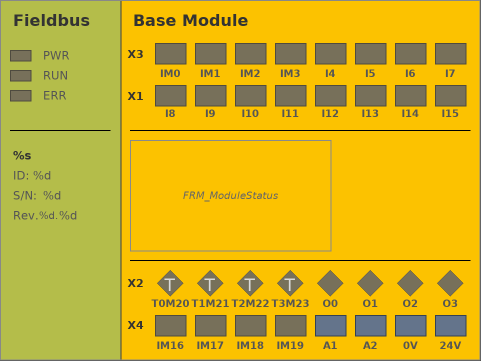
VISUALIZATION FRM_ModuleBase  // 481x361
VAR_IN_OUT
   stFieldbusData: ST_PNOZModuleData;
   stBaseModuleData: ST_PNOZModuleData;
END_VAR
    Rectangle (120,0 361x361)
    Frame (130,140 201x111)
        shows FRM_ModuleStatus(bPower := stBaseModuleData.stLEDState.bPower, bRun := stBaseModuleData.stLEDState.bRun, bDiag := stBaseModuleData.stLEDState.bDiag, bFault := stBaseModuleData.stLEDState.bFault, bInputFault := stBaseModuleData.stLEDState.bInputFault, bOutputFault := stBaseModuleData.stLEDState.bOutputFault, sName := stBaseModuleData.sName, nID := stBaseModuleData.nID, nSerialNumber := stBaseModuleData.nSerialNumber, anRevision := stBaseModuleData.anDeviceVersion)
    Line (130,130) (470,130)
    Line (130,260) (470,260)
    Label (120,44 31x21), "X3"
    Label (120,86 31x21), "X1"
    Label (120,273 31x21), "X2"
    Label (120,315 31x21), "X4"
    Label (130,0 141x41), "Base Module"
    Rectangle (0,0 121x361)
    Label (10,0 101x41), "Fieldbus"
    Rectangle (10,50 21x11), colour toggle: stFieldbusData.stLEDState.bPower
    Label (40,50 41x11), "PWR"
    Rectangle (10,70 21x11), colour toggle: stFieldbusData.stLEDState.bRun
    Label (40,70 41x11), "RUN"
    Rectangle (10,90 21x11), colour toggle: stFieldbusData.stLEDState.bFault
    Label (40,90 41x11), "ERR"
    Textfield (40,190 71x11), "%d", text variable: stFieldbusData.nSerialNumber
    Textfield (30,170 81x11), "%d", text variable: stFieldbusData.nID
    Textfield (10,150 101x11), "%s", text variable: stFieldbusData.sName
    Label (10,170 21x11), "ID:"
    Label (10,190 31x11), "S/N:"
    Line (10,130) (110,130)
    Rectangle (155,43 31x21), colour toggle: stBaseModuleData.anInput[1].b0
    Rectangle (195,43 31x21), colour toggle: stBaseModuleData.anInput[1].b1
    Rectangle (235,43 31x21), colour toggle: stBaseModuleData.anInput[1].b2
    Rectangle (275,43 31x21), colour toggle: stBaseModuleData.anInput[1].b3
    Rectangle (315,43 31x21), colour toggle: stBaseModuleData.anInput[1].b4
    Rectangle (355,43 31x21), colour toggle: stBaseModuleData.anInput[1].b5
    Rectangle (395,43 31x21), colour toggle: stBaseModuleData.anInput[1].b6
    Rectangle (435,43 31x21), colour toggle: stBaseModuleData.anInput[1].b7
    Label (150,68 41x11), "IM0"
    Label (190,68 41x11), "IM1"
    Label (230,68 41x11), "IM2"
    Label (270,68 41x11), "IM3"
    Label (310,68 41x11), "I4"
    Label (350,68 41x11), "I5"
    Label (390,68 41x11), "I6"
    Label (430,68 41x11), "I7"
    Rectangle (155,85 31x21), colour toggle: stBaseModuleData.anInput[2].b0
    Label (150,108 41x11), "I8"
    Label (190,108 41x11), "I9"
    Label (230,108 41x11), "I10"
    Label (270,108 41x11), "I11"
    Label (310,108 41x11), "I12"
    Label (350,108 41x11), "I13"
    Label (390,108 41x11), "I14"
    Label (430,108 41x11), "I15"
    Rectangle (195,85 31x21), colour toggle: stBaseModuleData.anInput[2].b1
    Rectangle (235,85 31x21), colour toggle: stBaseModuleData.anInput[2].b2
    Rectangle (275,85 31x21), colour toggle: stBaseModuleData.anInput[2].b3
    Rectangle (315,85 31x21), colour toggle: stBaseModuleData.anInput[2].b3
    Rectangle (355,85 31x21), colour toggle: stBaseModuleData.anInput[2].b5
    Rectangle (395,85 31x21), colour toggle: stBaseModuleData.anInput[2].b6
    Rectangle (435,85 31x21), colour toggle: stBaseModuleData.anInput[2].b7
    Polygon (157,283) (170,270) (183,283) (170,296) (170,296), colour toggle: stBaseModuleData.anOutput[2].b4
    Label (150,298 41x11), "T0M20"
    Label (190,298 41x11), "T1M21"
    Label (230,298 41x11), "T2M22"
    Label (270,298 41x11), "T3M23"
    Label (310,298 41x11), "O0"
    Label (350,298 41x11), "O1"
    Label (390,298 41x11), "O2"
    Label (430,298 41x11), "O3"
    Polygon (197,283) (210,270) (223,283) (210,296) (210,296), colour toggle: stBaseModuleData.anOutput[2].b5
    Polygon (237,283) (250,270) (263,283) (250,296) (250,296), colour toggle: stBaseModuleData.anOutput[2].b6
    Polygon (277,283) (290,270) (303,283) (290,296) (290,296), colour toggle: stBaseModuleData.anOutput[2].b7
    Polygon (317,283) (330,270) (343,283) (330,296) (330,296), colour toggle: stBaseModuleData.anOutput[1].b0
    Polygon (357,283) (370,270) (383,283) (370,296) (370,296), colour toggle: stBaseModuleData.anOutput[1].b1
    Polygon (397,283) (410,270) (423,283) (410,296) (410,296), colour toggle: stBaseModuleData.anOutput[1].b2
    Polygon (437,283) (450,270) (463,283) (450,296) (450,296), colour toggle: stBaseModuleData.anOutput[1].b3
    Rectangle (155,315 31x21), colour toggle: stBaseModuleData.anInput[3].b0
    Label (150,340 41x11), "IM16"
    Label (190,340 41x11), "IM17"
    Label (230,340 41x11), "IM18"
    Label (270,340 41x11), "IM19"
    Label (310,340 41x11), "A1"
    Label (350,340 41x11), "A2"
    Label (390,340 41x11), "0V"
    Label (430,340 41x11), "24V"
    Rectangle (195,315 31x21), colour toggle: stBaseModuleData.anInput[3].b1
    Rectangle (235,315 31x21), colour toggle: stBaseModuleData.anInput[3].b2
    Rectangle (275,315 31x21), colour toggle: stBaseModuleData.anInput[3].b3
    Rectangle (315,315 31x21)
    Rectangle (355,315 31x21)
    Rectangle (395,315 31x21)
    Rectangle (435,315 31x21)
    Label (157,275 26x20), "T"
    Label (197,275 26x20), "T"
    Label (237,275 26x20), "T"
    Label (277,275 26x20), "T"
    Textfield (40,210 21x11), "%d.", text variable: stFieldbusData.anDeviceVersion[1]
    Label (10,210 31x11), "Rev."
    Textfield (56,210 21x11), "%d", text variable: stFieldbusData.anDeviceVersion[2]
END_VISUALIZATION

(* stored: Version 1.1.0.1
   Visu FRM_ModuleBase: Id {12700075-affc-0e2a-1d48-8a87fd53542f} *)
